(* IEC 61131-3 sources: kns-port-domestic/tools/port_metrics_tests/fixtures/lib/src/POUs/FB_Base, 1 file *)

(* ---- FB_Base.decl.st ---- *)
FUNCTION_BLOCK FB_Base
VAR_OUTPUT
    xFault : BOOL;
END_VAR
